Fanuc KAREL source: kx00029.KL

PROGRAM KX00029
%STACKSIZE=65535
%PRIORITY=65535
VAR
I : INTEGER
J : INTEGER
B : BOOLEAN
F : FILE
S : STRING[80]
P : XYZWPR
BEGIN
I=1
END KX00029
